// TIA Portal V20 export
// export: Created 2026-10-19T18:05:47.5877685Z, ExportSetting WithDefaults, DisplayName Totally Integrated Automation Portal, DisplayVersion V20 Update 6, DisplayName TIA Portal Openness, DisplayVersion V20 Update 6, DisplayName TIA Portal Version Control Interface, DisplayVersion V20 Update 6, DisplayName SINAMICS Startdrive Advanced, DisplayVersion V20 SP1, DisplayName SINAMICS Startdrive G130, G150, S120, S150, SINAMICS MV, G220, S200, S210, DisplayVersion V20 SP1, DisplayName SINAMICS Startdrive G110M, G120, G120C, G120D, G120P, G115D, DisplayVersion V20 SP1, DisplayName STEP 7 Professional, DisplayVersion V20 Update 6, DisplayName STEP 7 Safety, DisplayVersion V20 Update 2, DisplayName WinCC Basic/Comfort/Advanced, DisplayVersion V20 Update 6, DisplayName WinCC Unified, DisplayVersion V20 Update 6
FUNCTION "FindStringField" : String   // FC19, SCL
{ S7_Optimized_Access := 'TRUE' }
VERSION : 0.1
// stored: AutoNumber true, IsIECCheckEnabled false, SetENOAutomatically false, UDAEnableTagReadback false
   VAR_INPUT
      FieldName : String;
      JsonStr : String;
   END_VAR
   VAR_TEMP
      searchStr : String;
      foundPos : Int;
      resultStr : String;
      quotePos1 : Int;
      quotePos2 : Int;
   END_VAR
BEGIN
   // Sets search pattern → ex: '"loadstate":'
   #searchStr := CONCAT(IN1 := '"', IN2 := #FieldName);
   #searchStr := CONCAT(IN1 := #searchStr, IN2 := '" :');

   // Search in JSON
   #foundPos := FIND(IN1 := #JsonStr, IN2 := #searchStr);

   IF #foundPos > 0 THEN
       // Finds first quote after field
       #quotePos1 := FIND(IN1 := MID(IN := #JsonStr, P := #foundPos + LEN(#searchStr), L := 20), IN2 := '"');

       IF #quotePos1 > 0 THEN
           // Finds second quote after the first
           #quotePos2 := FIND(
                              IN1 := MID(IN := #JsonStr, P := #foundPos + LEN(IN := #searchStr) + #quotePos1, L := 10),
                              IN2 := '"'
           );

           IF #quotePos2 > 0 THEN
               #resultStr := MID(
                                 IN := #JsonStr,
                                 P := #foundPos + LEN(#searchStr) + #quotePos1,
                                 L := #quotePos2 - 1
               );
               #FindStringField := #resultStr;
               RETURN;
           END_IF;
       END_IF;
   END_IF;

   // If not found, returns empty string
   #FindStringField := '';
END_FUNCTION
